(* IEC 61131-3 sources: SRCI_CLIENT_PLC/RobotLibrary/Library/POUs/Additional/MC_ReadCallSubprogramCyclic/Structures, 2 files *)

(* ---- ReadCallSubprogramCyclicOutCmd.st ---- *)
{attribute 'pack_mode' := '1'}
// -------------------------------------------------------------------------
//  SRCI Robot Library
// -------------------------------------------------------------------------
//
//  Object:      ReadCallSubprogramCyclicOutCmd
//  Author:      Thorsten Brach
//  Date:        2024-08-11
//
//  Description:
//
//
//  Copyright:
//    (C) 2024 Thorsten Brach. All rights reserved
//             Licensed under the MIT License.
//
//  Disclaimer:
//    This project is provided without any guarantee and can be used for
//    private and commercial purposes. Any use is at the user’s
//    own risk and responsibility.
//
// -------------------------------------------------------------------------
TYPE ReadCallSubprogramCyclicOutCmd :
STRUCT
  /// Cyclic input data of subprogram
  /// ST-FIX F179: size from RobotLibraryConstants.CYCLIC_SUB_PROGRAM_DATA_MAX
  Data : ARRAY[0..RobotLibraryConstants.CYCLIC_SUB_PROGRAM_DATA_MAX] OF BYTE;
END_STRUCT
END_TYPE

(* ---- ReadCallSubprogramCyclicParCmd.st ---- *)
{attribute 'pack_mode' := '1'}
// -------------------------------------------------------------------------
//  SRCI Robot Library
// -------------------------------------------------------------------------
//
//  Object:      UnitMeasurementParCmd
//  Author:      Thorsten Brach
//  Date:        2024-08-11
//
//  Description:
//
//
//  Copyright:
//    (C) 2024 Thorsten Brach. All rights reserved
//             Licensed under the MIT License.
//
//  Disclaimer:
//    This project is provided without any guarantee and can be used for
//    private and commercial purposes. Any use is at the user’s
//    own risk and responsibility.
//
// -------------------------------------------------------------------------
TYPE ReadCallSubprogramCyclicParCmd :
STRUCT
END_STRUCT
END_TYPE
